(* IEC 61131-3 sources: JingjiangArm/moonboxpro_arm_8.4/Application/Application/任务列表/ExtTask/动作处理/报警及提示, 6 files *)

(* ---- ENUM_MechanicalPart.st ---- *)
(*@CES
Name=ENUM_MechanicalPart
Type=Gvl
TypeGuid=2db5746d-d284-4425-9f7f-2663a34b0ebc
Guid=15e29af9-ac32-46fe-9cbd-84b481b11a74
HasDeclaration=True
HasImplementation=False
*)
{DECLARATION}
// {attribute 'qualified_only'}
// {attribute 'strict'}
TYPE ENUM_MechanicalPart :
(
	enum_member := 0,
	MECHANICALPART_PRNROLLER 	:= 3001,
	MECHANICALPART_NETROLLER 	:= 3002,
	MECHANICALPART_BOTTOMROLLER := 3003,
	MECHANICALPART_IF 			:= 3004,
	MECHANICALPART_OF 			:= 3005,
	MECHANICALPART_UW_A 		:= 3006,
	MECHANICALPART_UW_B 		:= 3007,
	MECHANICALPART_RW_A 		:= 3008,
	MECHANICALPART_RW_B 		:= 3009,
	MECHANICALPART_CENTERROLLER := 3010,
	MECHANICALPART_PRN_PRESS_M	:= 3011,
	MECHANICALPART_PRN_PRESS_G  := 3012,
	MECHANICALPART_NET_PRESS_M	:= 3013,
	MECHANICALPART_NET_PRESS_G  := 3014,
	MECHANICALPART_STR_PRESS_M	:= 3015,
	MECHANICALPART_STR_PRESS_G  := 3016,
	MECHANICALPART_INK_ROLLER	:= 3017,
	MECHANICALPART_SCRAPER		:= 3018,
	MECHANICALPART_HORZ			:= 3019,
	MECHANICALPART_PHOTOCELL	:= 3020

);
END_TYPE

	(*机械位置信息*)
(*
3001-----------------版辊
3002-----------------网辊
3003-----------------底辊
3004-----------------放牵
3005-----------------收牵
3006-----------------放料A
3007-----------------放料B
3008-----------------收料A
3009-----------------收料B
3010-----------------中心辊
3011-----------------版辊压力操作侧
3012-----------------版辊压力传动侧
3013-----------------网辊压力操作侧
3014-----------------网辊压力传动侧
3015-----------------张带压力操作侧
3016-----------------张带压力传动侧
3017-----------------递墨辊变频
3018-----------------刮刀变频
3019-----------------横向
3020-----------------光电眼
*)
{IMPLEMENTATION}

(* ---- StGetMotionSts.st ---- *)
(*@CES
Name=StGetMotionSts
Type=Gvl
TypeGuid=2db5746d-d284-4425-9f7f-2663a34b0ebc
Guid=76a34838-b972-4ac5-910f-8233101ca817
HasDeclaration=True
HasImplementation=False
*)
{DECLARATION}
TYPE StGetMotionSts :
STRUCT
	(*通过指令GT_RN_Getstaionsts获取*)
	uiVirtual_Cnt					: UINT;//虚拟码盘基数
	wVirtual_Sts: WORD;
	wNet_Status: WORD;
	wErr_a_Count: WORD;
	wErr_b_Count: WORD;
	wBreakCnt: WORD;
	wMotor_Temperature: WORD;
	wDriver_Temperature: WORD;
	wBus_Vol: WORD;
	(*通过指令GTN_GetDriverSts获取*)
	dwDriverSts: DWORD;
	(*通过指令GTN_GetServoAlarmInfo获取*)
	dwAlarmDetail: DWORD;
	(*通过大指令获取*)
	dwMotionSts: DWORD;
	lrPos_Prf: LREAL;
	lrPos_Enc: LREAL;
	lrVel_Prf: LREAL;
	lrVel_Enc: LREAL;
	lrPrfAcc: LREAL;//2026.5.8.112931新增

END_STRUCT
END_TYPE

{IMPLEMENTATION}

(* ---- StPTSts.st ---- *)
(*@CES
Name=StPTSts
Type=Gvl
TypeGuid=2db5746d-d284-4425-9f7f-2663a34b0ebc
Guid=280ed72c-8fcd-4475-a4e8-3c9693214690
HasDeclaration=True
HasImplementation=False
*)
{DECLARATION}
TYPE StPTSts :
STRUCT
	rtnSts:				INT;
	space:				INT;
	temperature:		INT;
	pfr:				DWORD;
	enc:				DWORD;
	vel:				INT;
	driverSts:			INT;
	driverErr:			INT;
	netPortSts:			INT;
	netRunSts:			INT;
	netPortErr_a:		INT;
	netPortErr_b:		INT;
	motionSts:			DWORD;
	modal:				WORD;
	virtualCnt:			WORD;
	virtualSts:			WORD;

	trigTime:			DWORD;
	trigCnt:			BYTE;
	brakeCnt:			WORD;
	driverCurrent:		WORD;
	driverTemp:			WORD;

	ai1_temp:			INT;
	ai2_temp:			INT;
	vdc:				INT;
	driverErr_high:		INT;
	sys_lock: 			DWORD;
	enc_lock:			DWORD;
	di:				WORD;

	rvsData_0:			WORD;
	encTemp:			WORD;
	rvsData_1:			WORD;
	rvsData_2:			DWORD;
	rvsData_3:			DWORD;
END_STRUCT
END_TYPE

{IMPLEMENTATION}

(* ---- KS_StationOnline.st ---- *)
(*@CES
Name=KS_StationOnline
Type=FunctionBlock
TypeGuid=6f9dac99-8de1-4efc-8465-68ac443b7d08
Guid=46162c4a-8077-432f-856c-536c68fec6ca
HasDeclaration=True
HasImplementation=True
*)
{DECLARATION}
FUNCTION KS_StationOnline : INT //2026.5.19.103428判断站点是否在线
VAR_INPUT
	i_iStationId: INT;
	i_pstStationInf_KS: POINTER TO StStationInfo_KS;
END_VAR
VAR
	iN: INT;
END_VAR

{IMPLEMENTATION}
KS_StationOnline:= 0;
IF i_iStationId>=0 AND i_iStationId<=MAX_STATION_NUM AND
	i_pstStationInf_KS<>0 THEN
	FOR iN:= 1 TO i_pstStationInf_KS^.iStationNum BY 1 DO
		IF i_pstStationInf_KS^.aiStationId_List[iN]= i_iStationId THEN
			KS_StationOnline:= 1;//返回只=1说明正常在线
			EXIT;
		END_IF
		IF iN= i_pstStationInf_KS^.iStationNum AND
			KS_StationOnline=0 THEN//离线
			KS_StationOnline:= -2;
		END_IF
	END_FOR
ELSE
	KS_StationOnline:= -1;
END_IF

(* ---- KS_FB_AlarmDisList.st ---- *)
(*@CES
Name=KS_FB_AlarmDisList
Type=FunctionBlock
TypeGuid=6f9dac99-8de1-4efc-8465-68ac443b7d08
Guid=9df2daeb-e031-42e6-924b-50f6708c13fd
HasDeclaration=True
HasImplementation=True
*)
{DECLARATION}
FUNCTION_BLOCK KS_FB_AlarmDisList
VAR_INPUT
	i_xEn:BOOL;
	i_iGrpId : INT;(*系ID*)
	i_iUnitNum:INT;
	i_pstStSysParam								: POINTER TO StSysParam;(*机器参数|*)
	i_pastStIOMap_Main_FE						: POINTER TO ARRAY [1..4] OF StIOMap_Main_FE;(*轴io数据区域|AB系*)
	i_pastStIOMap_Axis_FE					: POINTER TO ARRAY [1..MAX_UNIT_NUM] OF StIOMap_Axis_FE;(*轴io数据区域|*)
	i_pstStIOMap_Uw: POINTER TO StIOMap_UwRw_FE; (* 放料io|分A/B系 *)
	i_pstStIOMap_Rw: POINTER TO StIOMap_UwRw_FE; (* 收料io|分A/B系 *)
END_VAR
VAR_OUTPUT
	o_xEn:BOOL;
END_VAR
VAR
	iN : INT;
	iM : INT;
	iRtn : INT;
	iCustomerName: INT;
	afbRTrig_Estop:ARRAY [1..MAX_UNIT_NUM] OF R_TRIG;(*急停沿处理*)
	afbRTrig_Estop_UwRw:ARRAY [1..2] OF R_TRIG;(*收放料急停沿处理*)
	afbRTrig_Estop_IfOf:R_TRIG;(*收放料急停沿处理*)
	afbRTrig_PreStart: R_TRIG;(*预启动沿处理*)
	afbRTrig_Ink: R_TRIG;(*匀墨沿处理*)
	afbRTrig_Tension: R_TRIG;(*张力投入沿处理*)
	afbRTrig_Print: R_TRIG;(*印刷沿处理*)
	afbRTrig_Acc: R_TRIG;(*手动加速沿处理*)
	afbRTrig_Dec: R_TRIG;(*手动减速沿处理*)
	afbRTrig_Stop: R_TRIG;(*印刷沿处理*)
	xAxisInch_Print: BOOL;//点动2023.9.27.153613|收放牵|收放料|底辊|中心辊
	fbtrig_Inch_Print: R_TRIG;
	fbtrig_Inch_Stop: R_TRIG;
	fbtrig_Ink_Unit: R_TRIG;

	sAlarmMsg : STRING;
	sAlarmUnitId : STRING;
	iMsgId_Rec : INT := 1600;;
	iAlarmId_Rec : INT := 1600;
	iAlarm_TypeId_Rec : INT := 1600;

	afbRTrig_UnitPanel:ARRAY [1..MAX_UNIT_NUM,1..18] OF R_TRIG;(*收放料急停沿处理*)

	sAdjSts : STRING;
	sAlarmContent : STRING;
	(*2025.03.04.153303//网版电机开关沿处理*)
	afbtrig_NetMotorNo:ARRAY [1..MAX_UNIT_NUM] OF R_TRIG;
	afbtrig_NetMotorOff:ARRAY [1..MAX_UNIT_NUM] OF F_TRIG;
	(*2025.03.04.153303//走纸点动沿处理*)
	afbtrig_JogPaperNo:ARRAY [1..MAX_UNIT_NUM] OF R_TRIG;
	afbtrig_JogPaperOff:ARRAY [1..MAX_UNIT_NUM] OF F_TRIG;
END_VAR

{IMPLEMENTATION}
IF i_xEn THEN
	IF i_pstStSysParam <> 0 AND
		i_pstStSysParam <> 0 AND
		i_pastStIOMap_Main_FE <> 0 AND
		i_pastStIOMap_Axis_FE <> 0 AND
		i_pstStIOMap_Uw <> 0 AND
		i_pstStIOMap_Rw <> 0 THEN

		//收放料急停
		afbRTrig_Estop_UwRw[1](CLK:=i_pstStIOMap_Uw^.i_xEstop);
		afbRTrig_Estop_UwRw[2](CLK:=i_pstStIOMap_Rw^.i_xEstop);

		IF afbRTrig_Estop_UwRw[1].Q THEN
			//2026.1.20.140626 | + | 增加打印测试流程
			KS_HY_AddMsgToLog(g_pstStHYLogFifo, LOG_LEVEL_INFO, 'UW_EStop!', BOOL_TO_STRING(TRUE));
		END_IF
		IF afbRTrig_Estop_UwRw[2].Q THEN
			//2026.1.20.140626 | + | 增加打印测试流程
			KS_HY_AddMsgToLog(g_pstStHYLogFifo, LOG_LEVEL_INFO, 'RW_EStop!', BOOL_TO_STRING(TRUE));
		END_IF
		//牵引、界面急停
		afbRTrig_Estop_IfOf(CLK:=i_pastStIOMap_Main_FE^[1].i_xEstop OR i_pastStIOMap_Main_FE^[2].i_xEstop OR i_pastStIOMap_Main_FE^[3].i_xEstop OR i_pastStIOMap_Main_FE^[4].i_xEstop);
		IF afbRTrig_Estop_IfOf.Q THEN
			//2026.1.20.140626 | + | 增加打印测试流程
			KS_HY_AddMsgToLog(g_pstStHYLogFifo, LOG_LEVEL_INFO, 'IFOF_EStop!', BOOL_TO_STRING(TRUE));
		END_IF

		//预启动
		afbRTrig_PreStart(CLK:=i_pastStIOMap_Main_FE^[1].i_xPreStart OR i_pastStIOMap_Main_FE^[2].i_xPreStart OR i_pastStIOMap_Main_FE^[3].i_xPreStart OR i_pastStIOMap_Main_FE^[4].i_xPreStart);
		IF afbRTrig_PreStart.Q THEN
			//2026.1.20.140626 | + | 增加打印测试流程
			KS_HY_AddMsgToLog(g_pstStHYLogFifo, LOG_LEVEL_INFO, 'IFOF_PreStart!', BOOL_TO_STRING(TRUE));
		END_IF

		//匀墨
		afbRTrig_Ink(CLK:=i_pastStIOMap_Main_FE^[1].i_xInk OR i_pastStIOMap_Main_FE^[2].i_xInk OR i_pastStIOMap_Main_FE^[3].i_xInk OR i_pastStIOMap_Main_FE^[4].i_xInk);
		IF afbRTrig_Ink.Q THEN
			//2026.1.20.140626 | + | 增加打印测试流程
			KS_HY_AddMsgToLog(g_pstStHYLogFifo, LOG_LEVEL_INFO, 'IFOF_Ink!', BOOL_TO_STRING(TRUE));
		END_IF

		//张力投入
		afbRTrig_Tension(CLK:=i_pastStIOMap_Main_FE^[1].i_xTension OR i_pastStIOMap_Main_FE^[2].i_xTension OR i_pastStIOMap_Main_FE^[3].i_xTension OR i_pastStIOMap_Main_FE^[4].i_xTension);
		IF afbRTrig_Tension.Q THEN
			//2026.1.20.140626 | + | 增加打印测试流程
			KS_HY_AddMsgToLog(g_pstStHYLogFifo, LOG_LEVEL_INFO, 'IFOF_Tension!', BOOL_TO_STRING(TRUE));
		END_IF

		//印刷
		afbRTrig_Print(CLK:=i_pastStIOMap_Main_FE^[1].i_xPrint OR i_pastStIOMap_Main_FE^[2].i_xPrint OR i_pastStIOMap_Main_FE^[3].i_xPrint OR i_pastStIOMap_Main_FE^[4].i_xPrint);
		IF afbRTrig_Print.Q THEN
			//2026.1.20.140626 | + | 增加打印测试流程
			KS_HY_AddMsgToLog(g_pstStHYLogFifo, LOG_LEVEL_INFO, 'IFOF_Print!', BOOL_TO_STRING(TRUE));
		END_IF

		//加速
		afbRTrig_Acc(CLK:=i_pastStIOMap_Main_FE^[1].i_xAcc OR i_pastStIOMap_Main_FE^[2].i_xAcc OR i_pastStIOMap_Main_FE^[3].i_xAcc OR i_pastStIOMap_Main_FE^[4].i_xAcc);
		IF afbRTrig_Acc.Q THEN
			KS_HY_AddMsgToLog(g_pstStHYLogFifo, LOG_LEVEL_INFO, 'IFOF_Acc!', BOOL_TO_STRING(TRUE));
		END_IF

		//减速
		afbRTrig_Dec(CLK:=i_pastStIOMap_Main_FE^[1].i_xDec OR i_pastStIOMap_Main_FE^[2].i_xDec OR i_pastStIOMap_Main_FE^[3].i_xDec OR i_pastStIOMap_Main_FE^[4].i_xDec);
		IF afbRTrig_Dec.Q THEN
			KS_HY_AddMsgToLog(g_pstStHYLogFifo, LOG_LEVEL_INFO, 'IFOF_Dec!', BOOL_TO_STRING(TRUE));
		END_IF

		//停止
		afbRTrig_Stop(CLK:=i_pastStIOMap_Main_FE^[1].i_xStop OR i_pastStIOMap_Main_FE^[2].i_xStop OR i_pastStIOMap_Main_FE^[3].i_xStop OR i_pastStIOMap_Main_FE^[4].i_xStop);
		IF afbRTrig_Stop.Q THEN
			KS_HY_AddMsgToLog(g_pstStHYLogFifo, LOG_LEVEL_INFO, 'IFOF_Stop!', BOOL_TO_STRING(TRUE));
		END_IF

		//色组急停
		FOR iN:= 1 TO i_iUnitNum BY 1 DO
			//pstStUnitParam := ADR(i_pstStSysParam^.astStUnitParam[iN]);
			afbRTrig_Estop[iN](CLK:= i_pastStIOMap_Axis_FE^[iN].i_xEstop);
			IF afbRTrig_Estop[iN].Q THEN
				KS_HY_AddMsgToLog(g_pstStHYLogFifo, LOG_LEVEL_INFO, 'EStop Unit: ', INT_TO_STRING(iN));
			END_IF

			afbtrig_JogPaperNo[iN](CLK:= i_pastStIOMap_Axis_FE^[iN].i_xJogPaper);
			afbtrig_JogPaperOff[iN](CLK:= i_pastStIOMap_Axis_FE^[iN].i_xJogPaper);

			//走纸点动开关
			IF afbtrig_JogPaperNo[iN].Q THEN
				KS_HY_AddMsgToLog(g_pstStHYLogFifo, LOG_LEVEL_INFO, 'JogPaperOn Unit: ', INT_TO_STRING(iN));
			END_IF

			IF afbtrig_JogPaperOff[iN].Q THEN
				KS_HY_AddMsgToLog(g_pstStHYLogFifo, LOG_LEVEL_INFO, 'JogPaperOff Unit: ', INT_TO_STRING(iN));
			END_IF
		END_FOR

		IF iMsgId_Rec <> i_pstStSysParam^.astStGrpParam_UnSave[i_iGrpId].iPromptMsg OR iAlarm_TypeId_Rec <> i_pstStSysParam^.astStGrpParam_UnSave[i_iGrpId].iAlarm_TypeId OR
			iAlarmId_Rec <> i_pstStSysParam^.astStGrpParam_UnSave[i_iGrpId].iAlarm_UnitId THEN

			KS_HY_AddMsgToLog(g_pstStHYLogFifo, LOG_LEVEL_INFO, 'iPromptMsg: ', INT_TO_STRING(i_pstStSysParam^.astStGrpParam_UnSave[i_iGrpId].iPromptMsg));
			//KS_HY_AddMsgToLog(g_pstStHYLogFifo, LOG_LEVEL_INFO, 'iAlarm_TypeId: ', INT_TO_STRING(i_pstStSysParam^.astStGrpParam_UnSave[i_iGrpId].iAlarm_TypeId));
			KS_HY_AddMsgToLog(g_pstStHYLogFifo, LOG_LEVEL_INFO, 'iAlarm_UnitId: ', INT_TO_STRING(i_pstStSysParam^.astStGrpParam_UnSave[i_iGrpId].iAlarm_UnitId));
		END_IF
		iMsgId_Rec := i_pstStSysParam^.astStGrpParam_UnSave[i_iGrpId].iPromptMsg;
		iAlarmId_Rec := i_pstStSysParam^.astStGrpParam_UnSave[i_iGrpId].iAlarm_UnitId;
		iAlarm_TypeId_Rec := i_pstStSysParam^.astStGrpParam_UnSave[i_iGrpId].iAlarm_TypeId;

		//2025.01.04.111645 | 空转
		fbtrig_Ink_Unit(CLK:=g_axInk_Unit[1]);
		IF fbtrig_Ink_Unit.Q THEN
			KS_HY_AddMsgToLog(g_pstStHYLogFifo, LOG_LEVEL_INFO, 'Ink!', BOOL_TO_STRING(TRUE));
		END_IF
	END_IF
END_IF

(* ---- KS_FB_GrpFailureProc.st ---- *)
(*@CES
Name=KS_FB_GrpFailureProc
Type=FunctionBlock
TypeGuid=6f9dac99-8de1-4efc-8465-68ac443b7d08
Guid=09d385a5-873d-4de4-8b5b-a35479951d22
HasDeclaration=True
HasImplementation=True
*)
{DECLARATION}
FUNCTION_BLOCK KS_FB_GrpFailureProc
VAR_INPUT
	i_xEn: BOOL;
	i_iGrpId: INT;
	i_iCycle_Time: INT;
	i_byGrpUnitNum: INT;
	i_abyAxisList: ARRAY [1..MAX_UNIT_NUM] OF BYTE;
	i_iGrpAllStationNum: INT;
	i_aiStationList: ARRAY [1..MAX_STATION_NUM] OF INT;
	i_pstStSysParam: POINTER TO StSysParam;
	i_pastStGetMotionSts: POINTER TO ARRAY [1..MAX_STATION_NUM] OF StGetMotionSts;
	i_pastStAxisIdListInf :POINTER TO ARRAY [1..128] OF StAxisIdListInf;
	i_pastStIOMap_Main_FE	: POINTER TO ARRAY [1..4] OF StIOMap_Main_FE;(*轴io数据区域|*)
	i_pastStIOMap_AxisExtra: POINTER TO ARRAY [1..MAX_UNIT_NUM] OF StIOMap_Axis_Extra_FE;(*色组io|*)
	i_xLostPressure							: BOOL;(*气压低报警|不允许开机*)
	i_xPrnRollerLoose_AtLeast1				: BOOL;(*至少一色夹板松报警|不允许开机*)
	i_xbrakeResistanceTempHigh_AtLeast1		: BOOL;(*至少一色制动电阻温度高*)
	i_xHorzMotorAlarmAtLeastOne:BOOL;(*2022.6.28.000617*)
	i_xEstopBtnDne:BOOL;(*急停按下了|2022.6.28.150049*)
	i_xFlag_FastStopBtnDn: BOOL;
	i_xTowerInvAlarm_Uw:BOOL;(*2022.6.28.161545|来自altma特殊处理*)
	i_xTowerInvAlarm_Rw: BOOL;	(*  *)
	i_xInverterAlarmCurAxis_Uw				: BOOL;(*放料变频器当前轴报警*)
	i_xInverterAlarmCurAxis_Rw				: BOOL;(*收料变频器当前轴报警*)
	i_xInverterAlarmPreAxis_Uw				: BOOL;(*放料变频器预驱轴报警*)
	i_xInverterAlarmPreAxis_Rw				: BOOL;(*收料变频器预驱轴报警*)
	i_xInverterAlarm_If				: BOOL;(*放牵变频器报警*)
	i_xInverterAlarm_Of				: BOOL;(*收牵变频器报警*)

	i_xReflectSensorLoss					: BOOL;
	i_iMoveErrCode							: INT;(*初始化错误代码
												0-正常
												1-使能异常
												2-模态0设置异常
												3-模态1设置异常
												4-规划器启动异常
												5-PT模式设置异常
												6-伺服打开超时
												7-PT规划异常*)
	i_xAlarmHeating		: BOOL;
	i_xFlag_Alarm_LD:BOOL;
	i_pxFlag_Alarm_Rev_ErrorEnc:POINTER TO BOOL;(*编码器反转提示2022.9.16.135026*)
	i_iAxisId_Alarm_Rev:INT;(*编码器反转轴号*)
	i_xUwVolDiamMeasurementFailed: BOOL;
	i_dwAvailPhys_kB				: DWORD;(*有效的物理内存@小于一定阈值报警提示*)
	i_wAvailPhysAlarm_Kb			: WORD;(*物理内存报警值@小于这个值报警提示*)
	i_xCompensate_Phase_Stop		: BOOL;(*停机恢复相位提示*)
	i_xMemAllocFailed				: BOOL;(*内存申请失败*)
	i_xNeedRestartPlc				: BOOL;
	i_pstStGetPrm					:POINTER TO TMultiMcFunctionReadPrm;
	i_pstStSysStationInf			:POINTER TO StSysStationInf;
END_VAR
VAR_OUTPUT
	o_xEn: BOOL;
	o_iErNo									: INT;(*错误代码\-1:输入参数有误\|*)
	o_xInverterErrReset_Uw					: BOOL;
	o_xInverterErrReset_Rw					: BOOL;
	o_xAlarmStillOnline						: BOOL;(* 2022.3.15.125119/h/报警依然在线 |只有在列表中打印信息置位*)
	o_xClrAlarmSts							: BOOL;(*清除报警状态|用于外部变量的手动清除*)

END_VAR
VAR_IN_OUT
	io_byAutoBackUpSts:BYTE;(*SDCTL自动备份状态@=1 提示|=2 显示备份弹窗 *)
END_VAR
VAR
	iN: INT;
	iMsgId: INT;(*提示信息代码*)
	iAlarm_TypeId : INT;
	iAlarm_UnitId : INT;
	iAxisId: INT;
	iUnitId: INT;
	iTypeId: INT;
	iCoreId: INT;
	iGroupId : INT;
	axAlarmFlag: ARRAY [1..MAX_STATION_NUM] OF BOOL;
	xFaultInLinkageAxises: BOOL := FALSE;(*联动的轴里有错误|*)
	xFaultInIf: BOOL;
	abyAxisFailedCnt_ServoAlarm: ARRAY [1..MAX_STATION_NUM] OF BYTE := [MAX_STATION_NUM(0)];(*伺服报警|*)
	pstStUnitParam_Save: POINTER TO StUnitParam_Save;
	pstStUnitParam_UnSave: POINTER TO StUnitParam_UnSave;
	iTemp: INT;
	iBit: INT;
	fbTrigWillAutoPreCut_Uw:R_TRIG;
	fbTrigWillAutoPreCut_Rw:R_TRIG;
	xWillAutoMaticPreCut_Uw: BOOL;
	xWillAutoMaticPreCut_Rw: BOOL;
	iLinkageAxisNum: INT;
	iPromptMsg: INT;
	fbToF_UwVolDiamMeasurement: TON;
	alrBuff_Read: ARRAY [1..MAX_UNIT_NUM] OF LREAL;
	diReadCount: DINT;

	iRtn : INT;
	astStStationSts : ARRAY [1..MAX_STATION_NUM] OF StStationSts;
	abyStationList: ARRAY [1..MAX_STATION_NUM] OF BYTE;
	adiClock : ARRAY [1..MAX_STATION_NUM] OF DINT;
	stStSetPrm : TSetMultiMcFunctionPrm;
	alTime_Test: ARRAY [1..10] OF LTIME;

	iAdjAxisId : INT;
	iRead_UnitId : INT;

	iReadSts_Page : INT := 1;

	iReadDriverSts_Page : INT;

	adwDriverSts : ARRAY [1..MAX_STATION_NUM] OF DWORD;

	(*2025-12-10 by sjw 非阻塞大指令*)
	aFB_Get_StartMcMUltiFunction: ARRAY[1..2] OF GTMC_StartMcMultiFunction;
	axExecute: ARRAY [1..2] OF BOOL;
	axDoneGet: ARRAY[1..2] OF BOOL := [TRUE, TRUE];
	axBusyGet: ARRAY[1..2] OF BOOL;
	axErrorGet: ARRAY[1..2] OF BOOL;
	aiErrorIdGet: ARRAY[1..2] OF INT;

	//2025.11.03.103620 | bai.zy | TEST_1103
	apData : ARRAY [1..MAX_UNIT_NUM] OF UINT;

	atiTimeReadWatch : ARRAY [1..MAX_UNIT_NUM] OF LTIME;

	iReadVirtualSts_UnitId : INT;

	alrBuff_Read2: ARRAY [1..MAX_UNIT_NUM,1..50] OF LREAL;

	adiReadCount: ARRAY [1..MAX_UNIT_NUM] OF DINT;
	iK : INT;

	//altime : ARRAY [1..20] OF LTIME;

	iCountRes : INT;
	iCurrentNum_Start : INT;
	iCurrentNum_End : INT;

	//2026.02.04.170811 | + | 这里需要把方向处理一下，只有主从轴的方向不一致才需要把从轴方向改了
	axGantryAxisIsRev : ARRAY [1..20,1..2] OF BOOL;//最大20组龙门，每组龙门两个轴
	iGantryAxisCount : INT;

	iUpdateEncPosStart : INT;
	iUpdateEncPosEnd : INT;

	iGetDriverStsAxis : INT;
	iGetStsCnt : INT;
END_VAR

{IMPLEMENTATION}
o_xEn:= i_xEn;
o_iErNo:= 0;
o_xAlarmStillOnline:= FALSE;(* 2022.3.15.125148/h/+ *)
o_xAlarmStillOnline:= FALSE;(* 2022.3.15.125148/h/+ *)
IF i_xEn THEN
	IF (i_iGrpId=1 OR i_iGrpId=2) AND
		i_byGrpUnitNum>=1 AND i_byGrpUnitNum<=MAX_UNIT_NUM AND
		i_pstStSysParam<>0 THEN
		IF i_iCycle_Time=0 THEN
			i_iCycle_Time:= gc_EXT_TSK_CYCLE_TIME;
		END_IF
		FOR iN:=1 TO i_iGrpAllStationNum BY 1 DO
// 			KS_HY_GetAxisIdForMotByStation(
// 				i_aiStationList[iN],
// 				ADR(iAxisId),
// 				ADR(iTypeId),
// 				ADR(iUnitId),
// 				ADR(iCoreId),
// 				ADR(iGroupId),
// 				ADR(iAdjAxisId),
// 				i_pastStAxisIdListInf
//				);
			KS_GetAxisIdForMotByStation_V2(
					i_iStationId:= i_aiStationList[iN],
					i_piAxisId:= ADR(iAxisId),
					i_piTypeId:= ADR(iTypeId),
					i_piUnitId:= ADR(iUnitId),
					i_piCoreId:= ADR(iCoreId),
					i_piGroupId:= ADR(iGroupId),
					i_piAdjAxisId:= ADR(iAdjAxisId),
					i_pstStSysStationInf:= i_pstStSysStationInf);
			(*报警处理*)
			IF NOT o_xClrAlarmSts THEN
				IF i_pastStGetMotionSts^[(iCoreId-1)* gc_ResCount_Profile +iAxisId].dwMotionSts.1 THEN(*bit1:报警*)
					IF abyAxisFailedCnt_ServoAlarm[iN]>5 THEN(*超过5个周期确定报警*)
//处理报警标志位
						axAlarmFlag[iN]:= TRUE;
					ELSE
						abyAxisFailedCnt_ServoAlarm[iN]:= abyAxisFailedCnt_ServoAlarm[iN]+1;
					END_IF
				ELSE
					abyAxisFailedCnt_ServoAlarm[iN]:= 0;
					IF axAlarmFlag[iN] THEN
						axAlarmFlag[iN]:= FALSE;
					END_IF
				END_IF
			END_IF
			Action_SysAlarmFlag();//报警标志赋值到全局变量
			o_xAlarmStillOnline:= o_xAlarmStillOnline OR axAlarmFlag[iN];
		END_FOR
		xFaultInLinkageAxises:= FALSE;
		FOR iN:=1 TO i_byGrpUnitNum BY 1 DO
			iUnitId:= i_abyAxisList[iN];
			pstStUnitParam_Save:= ADR(i_pstStSysParam^.astStUnitParam_Save[iUnitId]);
			pstStUnitParam_UnSave:= ADR(i_pstStSysParam^.astStUnitParam_UnSave[iUnitId]);
			IF NOT pstStUnitParam_Save^.xLinkage THEN
				;
			ELSE
				IF pstStUnitParam_UnSave^.xAxisAlarm_PrnRoller OR
					pstStUnitParam_UnSave^.xAxisAlarm_NetRoller OR
					pstStUnitParam_UnSave^.xAxisAlarm_BottomRoller OR
					pstStUnitParam_UnSave^.xAxisAlarm_Horz OR
					pstStUnitParam_UnSave^.xAxisAlarm_Prn_Pressure_M OR
					pstStUnitParam_UnSave^.xAxisAlarm_Prn_Pressure_G OR
					pstStUnitParam_UnSave^.xAxisAlarm_Net_Pressure_M OR
					pstStUnitParam_UnSave^.xAxisAlarm_Net_Pressure_G OR
					pstStUnitParam_UnSave^.xAxisAlarm_Str_Pressure_M OR
					pstStUnitParam_UnSave^.xAxisAlarm_Str_Pressure_G THEN
					(*色组内任意部位报警都当作急停处理吧*)
					(*but:压力电机报警可能不能急停？柔印时候再考虑一下*)
					IF NOT xFaultInLinkageAxises THEN
						xFaultInLinkageAxises:= TRUE;
					END_IF
				END_IF
			END_IF
		END_FOR
		(*上面处理了色组报警-同时收放料收放牵也要处理*)
		IF i_pstStSysParam^.astStGrpParam_UnSave[i_iGrpId].xAxisAlarm_CENTRAL OR
			i_pstStSysParam^.astStGrpParam_UnSave[i_iGrpId].xAxisAlarm_If OR
			i_pstStSysParam^.astStGrpParam_UnSave[i_iGrpId].xAxisAlarm_Of OR
			i_pstStSysParam^.astStGrpParam_UnSave[i_iGrpId].xAxisAlarm_Uw_A OR
			i_pstStSysParam^.astStGrpParam_UnSave[i_iGrpId].xAxisAlarm_Uw_B OR
			i_pstStSysParam^.astStGrpParam_UnSave[i_iGrpId].xAxisAlarm_Rw_A OR
			i_pstStSysParam^.astStGrpParam_UnSave[i_iGrpId].xAxisAlarm_Rw_B THEN
			IF NOT xFaultInLinkageAxises THEN
				xFaultInLinkageAxises:= TRUE;
			END_IF
		END_IF
		i_pstStSysParam^.astStGrpParam_UnSave[i_iGrpId].xFlag_LinkageAxisAlarm:= xFaultInLinkageAxises;
		(*到这里报警先处理完成了-下面处理提示信息*)
		(*是否出现报警再执行读取报警信息小指令？？先按每个周期都读吧*)
		iMsgId:= 0;
		iAlarm_TypeId := 0;
		iAlarm_UnitId := 0;
		Action_Msg_Alarm();
		Action_Msg_Tip();
		i_pstStSysParam^.astStGrpParam_UnSave[i_iGrpId].iPromptMsg:= iMsgId;
		i_pstStSysParam^.astStGrpParam_UnSave[i_iGrpId].iAlarm_TypeId:= iAlarm_TypeId;
		i_pstStSysParam^.astStGrpParam_UnSave[i_iGrpId].iAlarm_UnitId:= iAlarm_UnitId;
(*到这里就结束了-下面需要增加复位逻辑和读取状态逻辑*)
		Action_Alarm_ClearAndReset();
		Action_GrpGetMotionSts();
	END_IF
ELSE;
END_IF
